// TIA Portal V21 export
// export: Created 2026-11-11T00:47:27.1418872Z, ExportSetting WithDefaults, DisplayName Totally Integrated Automation Portal, DisplayVersion V21 Update 3, DisplayName STEP 7 Professional, DisplayVersion V21 Update 3, DisplayName STEP 7 Safety, DisplayVersion V21, DisplayName Tech WebApplication, DisplayVersion V21, DisplayName WinCC Basic/Comfort/Advanced, DisplayVersion V21 Update 3, DisplayName WinCC Unified, DisplayVersion V21 Update 3
FUNCTION_BLOCK "FB_Fbd_ex105"   // FB117, FBD
{ S7_Optimized_Access := 'TRUE' }
VERSION : 0.1
// stored: AutoNumber true, IsIECCheckEnabled false, IsRetainMemResEnabled false, MemoryReserve 100, SetENOAutomatically false, UDAEnableTagReadback false
   VAR_INPUT
      v_ob_nr : OB_TOD;
      v_sdt : DTL;
      v_local : Bool;
      v_period : Word;
      v_activate : Bool;
   END_VAR
   VAR_OUTPUT
      v_ret_val : Int;
   END_VAR
BEGIN

REGION Network 1: SET_TINTL - Set time-of-day interrupt
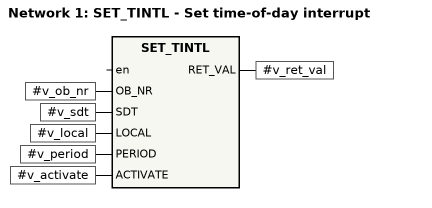
   #v_ret_val := SET_TINTL(OB_NR := #v_ob_nr,
                           SDT := #v_sdt,
                           LOCAL := #v_local,
                           PERIOD := #v_period,
                           ACTIVATE := #v_activate);
END_REGION
END_FUNCTION_BLOCK
